{attribute 'qualified_only'}
{attribute 'strict'}
{attribute 'to_string'}
TYPE E_AxisHomeSource : (
    Unknown := 0,
    NC := 1,
    Drive := 2
);
END_TYPE

(* stored: Version 1.1.0.1, ProductVersion 3.1.4026.20
   DUT E_AxisHomeSource: Id {2fa0fa69-546c-5566-ab5e-59ad7b2f8900} *)
